(* IEC 61131-3 sources: STAR-PLC-Agent/results/raw/codex_matrix_resume_20261114/codex_deepseek/PUB012/generation/compiler_records/compile_01, 1 file *)

(* ---- FB_Task.st ---- *)
FUNCTION_BLOCK FB_Task
VAR_INPUT
    THICKNESS_FAULT : BOOL;
    THICKNESS_SIGNAL_VALID : BOOL;
    CUTTING_RUN : BOOL;
    FaultTimestamp : DINT;
    CycleTime : TIME;
END_VAR
VAR_OUTPUT
    THICKNESS_ALARM : BOOL;
    Slab_Fault_Counter : UINT;
    Slab_Runtime_Accumulator : LTIME;
    Slab_Fault_History : ARRAY[0..4] OF DINT;
END_VAR
VAR
    _PrevValidFault : BOOL;
    _HoldActive : BOOL;
    _HoldTimer : TON;
    _FaultRise : BOOL;
END_VAR

_FaultRise := THICKNESS_SIGNAL_VALID AND THICKNESS_FAULT AND NOT _PrevValidFault;

IF NOT THICKNESS_SIGNAL_VALID THEN
    _HoldActive := FALSE;
    _HoldTimer(IN := FALSE, PT := T#500MS);
    THICKNESS_ALARM := FALSE;
ELSE
    IF _FaultRise THEN
        _HoldActive := TRUE;
        _HoldTimer(IN := FALSE, PT := T#500MS);
        _HoldTimer(IN := TRUE, PT := T#500MS);
    ELSE
        _HoldTimer(IN := _HoldActive, PT := T#500MS);
        IF _HoldTimer.Q THEN
            _HoldActive := FALSE;
        END_IF;
    END_IF;

    THICKNESS_ALARM := THICKNESS_FAULT OR _HoldActive;
END_IF;

IF _FaultRise THEN
    Slab_Fault_History[4] := Slab_Fault_History[3];
    Slab_Fault_History[3] := Slab_Fault_History[2];
    Slab_Fault_History[2] := Slab_Fault_History[1];
    Slab_Fault_History[1] := Slab_Fault_History[0];
    Slab_Fault_History[0] := FaultTimestamp;
    Slab_Fault_Counter := Slab_Fault_Counter + 1;
END_IF;

IF THICKNESS_SIGNAL_VALID AND NOT THICKNESS_FAULT AND CUTTING_RUN THEN
    Slab_Runtime_Accumulator := Slab_Runtime_Accumulator + TIME_TO_LTIME(CycleTime);
END_IF;

_PrevValidFault := THICKNESS_SIGNAL_VALID AND THICKNESS_FAULT;
END_FUNCTION_BLOCK
